(* CODESYS project maincontrol.library
   DefaultNamespace: KOSTAL.AF2024.Core.MainControl
   DocFormat: reStructuredText
   Description: Base Class of Machnie Main Control with 
      Cell_EXT using the ListOfInterface library instead of the generic array.
      The handler for the subscribers/stations is provided as well.
   Author: Frank Dümpelmann
   Title: KOSTAL.AF2024.Core.MainControl
   Version: 1.0.0.0
   Company: KOSTAL GmbH & Co.KG
   Placeholder: KOSTAL.AF2024.Core.MainControl

Project tree, tasks and I/O mapping:
  libraries: KOSTAL.AF2024.Core.functionResponse, 1.0.0.0 (KOSTAL GmbH & Co.KG); KOSTAL.AF2024.Core.ID, 1.0.0.0 (KOSTAL GmbH & Co.KG); KOSTAL.AF2024.Core.ListOf, 1.0.0.0 (KOSTAL GmbH & Co.KG); KOSTAL.AF2024.Core.Process, 1.0.0.0 (KOSTAL GmbH & Co.KG); KOSTAL.AF2024.Core.Settings, 1.0.0.0 (KOSTAL GmbH & Co.KG); KOSTAL.AF2024.Core.StringTools, 1.0.0.0 (KOSTAL GmbH & Co.KG); KOSTAL.AF2024.Core.System, 1.0.0.0 (KOSTAL GmbH & Co.KG)
  MainControl/
    Participant/
      ListOf/
        function block FB_ListOfParticipant [ST]: _setResult, _verifyMember, AddMember, Clear, Get_Member, IsValidParticipant, NumberOfMember, RegKey, RemoveMember, RemoveMemberByNumber
        interface I_ListOfParticipant: NumberOfMember, RegKey
        interface I_ListOfParticipant_Owner: AddMember, Clear, Get_Member, IsValidParticipant, NumberOfMember, RegKey, RemoveMember, RemoveMemberByNumber
      function block FB_Participant [ST]: FB_init, _clearRegisterInformation, Register, ParticipantName, Condition, Demand, ID, Linked, Mode, State
      interface I_Participant: Demand, ID, Mode, Register, Condition, ParticipantName, State, Linked
    function block FB_MainControl [ST]: _all_ErrorFree, _all_Finish, _all_Home, _all_OnToHome, _all_PowerOff, _all_PowerOn, _all_Run, _getNameAndID, _setResult, FB_exit, FB_init, Register, Unregister, condition, Demand, Device_ID, enableStopMode, ID, ID_RO, Mode, Participants, RunEmpty, step
    interface I_MainControl: condition, Demand, Device_ID, enableStopMode, ID_RO, Mode, Participants, RunEmpty, step
  MainControlState/
    interface I_T_MainControlState: CopyTo, Home, OnToHome, PowerOff, PowerOn, Run, RunToHome
    interface I_T_MainControlState_CopyFrom: CopyFrom
    interface I_T_MainControlState_Owner: clear, CopyFrom, CopyTo, Home, OnToHome, PowerOff, PowerOn, Run, RunToHome, SetUnique_Home, SetUnique_OnToHome, SetUnique_PowerOff, SetUnique_PowerOn, SetUnique_Run, SetUnique_RunToHome
    function block T_MainControlState [ST]: _clear_state, clear, CopyFrom, CopyTo, Home, OnToHome, PowerOff, PowerOn, Run, RunToHome, SetUnique_Home, SetUnique_OnToHome, SetUnique_PowerOff, SetUnique_PowerOn, SetUnique_Run, SetUnique_RunToHome
  ParticipantState/
    interface I_T_ParticipantState: Busy, CopyTo, Finish, Home, OnToHome, PowerOff, PowerOn
    interface I_T_ParticipantState_CopyFrom: CopyFrom
    interface I_T_ParticipantState_Owner: Busy, clear, CopyFrom, CopyTo, Finish, Home, OnToHome, PowerOff, PowerOn, SetUnique_Busy, SetUnique_Finish, SetUnique_Home, SetUnique_OnToHome, SetUnique_PowerOff, SetUnique_PowerOn
    function block T_ParticipantState [ST]: _clear_state, Busy, clear, CopyFrom, CopyTo, Finish, Home, OnToHome, PowerOff, PowerOn, SetUnique_Busy, SetUnique_Finish, SetUnique_Home, SetUnique_OnToHome, SetUnique_PowerOff, SetUnique_PowerOn
  Project Information/
    function F_GetCompany [ST]
    function F_GetTitle [ST]
    function F_GetVersion [ST]
  Version/
    global variables Global_Version
*)

// Version/Global_Version
{attribute 'TcGenerated'}
{attribute 'no-analysis'}
{attribute 'linkalways'}
// This function has been automatically generated from the project information.
VAR_GLOBAL CONSTANT
	{attribute 'const_non_replaced'}
	stLibVersion_KOSTAL_AF2024_Core_MainControl : ST_LibVersion := (iMajor := 1, iMinor := 0, iBuild := 0, iRevision := 0, nFlags := 0, sVersion := '1.0.0.0');
END_VAR

// MainControl/Participant/ListOf/FB_ListOfParticipant
(*
Extends the generic class with typed content.
*)
FUNCTION_BLOCK FB_ListOfParticipant EXTENDS KOSTAL_AF2024_Core_ListOf._FB_Interface_Base IMPLEMENTS I_ListOfParticipant, I_ListOfParticipant_Owner

VAR
	_PH_ID				: KOSTAL_AF2024_Core_ID.T_ID;	//placeholder for interfaces
	_PH_Condition 		: KOSTAL_AF2024_Core_Process.FB_processCondition;	//placeholder for interfaces
	_PH_State		 	: T_ParticipantState;	//placeholder for interfaces
	_PH_MainControlDemand		: T_MainControlState;	//placeholder for interfaces
	_PH_MainControlMode 		: KOSTAL_AF2024_Core_Process.T_processMode;	//placeholder for interfaces

	_Dummy	:	FB_Participant(ID:= _PH_ID, Condition:= _PH_Condition, State:= _PH_State);
END_VAR

METHOD PROTECTED _setResult
VAR_INPUT
	Status	: KOSTAL_AF2024_Core_Settings.T_MaxString;
	Success	: BOOL;
	Result	: KOSTAL_AF2024_Core_functionResponse.I_T_functionResponse_Owner;
END_VAR

IF Result = 0 THEN RETURN;	END_IF

Result.status:= Status;
Result.success:= Success;
END_METHOD

(*
	integrate here the veryfing of your interface type 
	only if verifing is passed [_verifyMember:= TRUE] the called metode will proceeded 
*)
METHOD PROTECTED _verifyMember : BOOL

VAR_INPUT
	Member	: KOSTAL_AF2024_Core_System.I_Interface;
	Result	: KOSTAL_AF2024_Core_functionResponse.I_T_functionResponse_Owner;
END_VAR

VAR
	_obj	: I_Participant;
	_bResult: BOOL;
END_VAR

_verifyMember:= SUPER^._verifyMember(Member, Result);

IF NOT _verifyMember THEN RETURN;	END_IF

//if member is I_participant?
_bResult:= __QUERYINTERFACE(Member, _obj);

IF NOT _bResult OR (_obj = 0) THEN
	IF Result <> 0 THEN
		Result.success:= FALSE;
		Result.status:= "no valid interface found";	
	END_IF	
	RETURN;
END_IF

//if 
IF NOT IsValidParticipant(_obj, Result)	THEN RETURN;	END_IF

_verifyMember:= TRUE;
END_METHOD

(*
	add new {Member} to end of list
*)
METHOD PUBLIC AddMember : BOOL

VAR_INPUT
	Member	: KOSTAL_AF2024_Core_System.I_Interface;
	Result	: KOSTAL_AF2024_Core_functionResponse.I_T_functionResponse_Owner;
END_VAR

AddMember:= SUPER^._addMember(Member, Result);

IF AddMember THEN	AddMember:= SUPER^._checkConsistency(Result);	END_IF
END_METHOD

//Clear the whole content
METHOD PUBLIC Clear

SUPER^._clear();
END_METHOD

METHOD PUBLIC Get_Member : I_Participant
VAR_INPUT
	Number		: UDINT;	//Participant which shall return
	Response	: KOSTAL_AF2024_Core_functionResponse.I_T_functionResponse_Owner;
END_VAR

VAR
	_Response	: KOSTAL_AF2024_Core_functionResponse.T_functionResponse;
	_Member			:	KOSTAL_AF2024_Core_System.I_Interface; 
	_obj			: I_Participant;
	_bResult	: BOOL;
	_found		: BOOL;
END_VAR
Get_Member:= _Dummy;

IF Number = 0 THEN
	IF Response <> 0 THEN	
		Response.success:= FALSE;	Response.status:= "Number is out of range";	
	END_IF
	RETURN;
END_IF

_found := _findMemberByIndex(Number - 1, _Member, _Response);
 
IF NOT _found OR NOT _Response.success THEN
 IF Response <> 0 THEN 
	Response.CopyFrom(_Response);	
	END_IF
 RETURN;
END_IF

_bResult:= __QUERYINTERFACE(_Member, _obj);

IF NOT _bResult THEN
	_Response.success:= FALSE;	_Response.status:= "__QUERYINTERFACE (I_RO) failed";
	IF Response <> 0 THEN 
		Response.CopyFrom(_Response);		
		END_IF
	RETURN;
END_IF

_Response.success:= TRUE;	_Response.status:= "Successful";
IF Response <> 0 THEN 
	Response.CopyFrom(_Response);	
END_IF

Get_Member:= _obj;
END_METHOD

METHOD PUBLIC IsValidParticipant : BOOL
VAR_INPUT
	Participant	: I_Participant;
	Result			: KOSTAL_AF2024_Core_functionResponse.I_T_functionResponse_Owner;
END_VAR

VAR
	_oParticipant 				: I_Participant;
	_bResult			: BOOL;
END_VAR
IsValidParticipant:= FALSE;

IF	Participant = 0 THEN	_setResult("no valid I_Participant INTERFACE", FALSE, Result);	RETURN; END_IF	

_bResult:= __QUERYINTERFACE( Participant, _oParticipant);

IF NOT _bResult 									THEN	_setResult("no valid I_Participant INTERFACE", FALSE, Result);	
ELSIF	_oParticipant = 0 									THEN	_setResult("no valid I_Participant INTERFACE", FALSE, Result);	
ELSIF	Participant = 0 						THEN	_setResult("no valid I_Participant INTERFACE", FALSE, Result);	
ELSIF Participant.Demand = 0	THEN	_setResult("no valid MainControlDemand INTERFACE", FALSE, Result);	
ELSIF Participant.Mode = 0		THEN	_setResult("no valid Mode INTERFACE", FALSE, Result);	
ELSIF Participant.Condition = 0		THEN	_setResult("no valid Condition INTERFACE", FALSE, Result);	
ELSIF Participant.ID = 0					THEN	_setResult("no valid ID INTERFACE", FALSE, Result);	
ELSIF Participant.State = 0				THEN	_setResult("no valid State INTERFACE", FALSE, Result);	
ELSE	IsValidParticipant:= TRUE;
END_IF
END_METHOD

//return the nnumber of items in List
PROPERTY PUBLIC NumberOfMember : UDINT
GET

NumberOfMember:= _NumberOfMember;
END_GET
END_PROPERTY

PROPERTY PUBLIC RegKey : UDINT
GET

RegKey:= _RegKey;
END_GET
END_PROPERTY

(*
	remove given {Member} from List
*)
METHOD PUBLIC RemoveMember : BOOL
VAR_INPUT
	Member	: KOSTAL_AF2024_Core_System.I_Interface;
	Result	: KOSTAL_AF2024_Core_functionResponse.I_T_functionResponse_Owner;
END_VAR

IF NOT _verifyMember(Member, Result) THEN	RETURN;	END_IF

RemoveMember:= _removeMember(Member, Result);

IF RemoveMember THEN	RemoveMember:= SUPER^._checkConsistency(Result);	END_IF
END_METHOD

(*
	remove given {Number} from List
*)
METHOD PUBLIC RemoveMemberByNumber : BOOL
VAR_INPUT
	Number	: UDINT;	//Position which shall deleted
	Result	: KOSTAL_AF2024_Core_functionResponse.I_T_functionResponse_Owner;
END_VAR
IF Number = 0 THEN
	IF Result <> 0  THEN
		Result.success:= FALSE;	
		Result.status:= "Number is out of range";	
	END_IF
	RETURN;
END_IF

RemoveMemberByNumber:= _removeMemberByIndex(Number - 1, Result);

IF RemoveMemberByNumber THEN	RemoveMemberByNumber:= SUPER^._checkConsistency(Result);	END_IF
END_METHOD

END_FUNCTION_BLOCK

// MainControl/Participant/ListOf/I_ListOfParticipant
(*
	Read-Only access to List
*)
INTERFACE I_ListOfParticipant EXTENDS KOSTAL_AF2024_Core_ListOf._I_Interface_Base

PROPERTY PUBLIC NumberOfMember : UDINT
GET
END_GET
END_PROPERTY

PROPERTY PUBLIC RegKey : UDINT
GET
END_GET
END_PROPERTY

END_INTERFACE

// MainControl/Participant/ListOf/I_ListOfParticipant_Owner
(*
	full access to List
*)
INTERFACE I_ListOfParticipant_Owner EXTENDS KOSTAL_AF2024_Core_ListOf._I_Interface_Base_Owner

(*
	add new {Member} to end of list
*)
METHOD PUBLIC AddMember : BOOL

VAR_INPUT
	Member	: KOSTAL_AF2024_Core_System.I_Interface;
	Result	: KOSTAL_AF2024_Core_functionResponse.I_T_functionResponse_Owner;
END_VAR
END_METHOD

//Clear the whole content
METHOD PUBLIC Clear
END_METHOD

METHOD PUBLIC Get_Member : I_Participant
VAR_INPUT
	Number		: UDINT;	//Participant which shall return
	Response	: KOSTAL_AF2024_Core_functionResponse.I_T_functionResponse_Owner;
END_VAR
END_METHOD

METHOD PUBLIC IsValidParticipant : BOOL
VAR_INPUT
	Participant	: I_Participant;
	Result			: KOSTAL_AF2024_Core_functionResponse.I_T_functionResponse_Owner;
END_VAR
END_METHOD

//return the nnumber of items in List
PROPERTY PUBLIC NumberOfMember : UDINT
GET
END_GET
END_PROPERTY

PROPERTY PUBLIC RegKey : UDINT
GET
END_GET
END_PROPERTY

(*
	remove given {Member} from List
*)
METHOD PUBLIC RemoveMember : BOOL
VAR_INPUT
	Member	: KOSTAL_AF2024_Core_System.I_Interface;
	Result	: KOSTAL_AF2024_Core_functionResponse.I_T_functionResponse_Owner;
END_VAR
END_METHOD

(*
	remove given {Number} from List
*)
METHOD PUBLIC RemoveMemberByNumber : BOOL
VAR_INPUT
	Number	: UDINT;	//Position which shall deleted
	Result	: KOSTAL_AF2024_Core_functionResponse.I_T_functionResponse_Owner;
END_VAR
END_METHOD

END_INTERFACE

// MainControl/Participant/I_Participant
(*

:Author: Frank Dümpelmann <f.duempelmann@kostal.com>, Martin Hundt <m.hundt@kostal.com>
:Date: 2018-10-29

Function
========
Interface for communication between stations and MainControl

Usage notes
===============
| All stations must be implemented with this interface



*)

INTERFACE I_Participant EXTENDS KOSTAL_AF2024_Core_System.I_Interface

(*State requirement for the participant*)
PROPERTY Demand : I_T_MainControlState
GET
END_GET
END_PROPERTY

(*
	ID of the participant
	{name} will handeld by participant
	{key} will handled by MainControl. 
*)
PROPERTY ID : KOSTAL_AF2024_Core_ID.I_T_ID
GET
END_GET
END_PROPERTY

(*Mode information for the participant*)
PROPERTY Mode : KOSTAL_AF2024_Core_process.I_T_processMode
GET
END_GET
END_PROPERTY

(*
	Called by MainControl
*)
METHOD PUBLIC Register
VAR_INPUT
	MainControlDemand	: I_T_MainControlState;
	MainControlMode		: KOSTAL_AF2024_Core_process.I_T_processMode;
	RegKey			: UDINT;
	Linked			: BOOL;
END_VAR
END_METHOD

(*Condition of the participant*)
PROPERTY Condition : KOSTAL_AF2024_Core_process.I_processCondition
GET
END_GET
END_PROPERTY

PROPERTY PUBLIC ParticipantName : KOSTAL_AF2024_Core_Settings.T_MaxString
GET
END_GET
END_PROPERTY

(*State of the participant*)
PROPERTY State : I_T_ParticipantState
GET
END_GET
END_PROPERTY

PROPERTY PUBLIC Linked : BOOL
GET
END_GET
END_PROPERTY

END_INTERFACE

// MainControlState/I_T_MainControlState
INTERFACE I_T_MainControlState EXTENDS KOSTAL_AF2024_Core_System.I_Interface

METHOD PUBLIC CopyTo
VAR_INPUT
	IN	:	I_T_MainControlState_CopyFrom;
END_VAR
END_METHOD

PROPERTY PUBLIC Home : BOOL
GET
END_GET
END_PROPERTY

PROPERTY PUBLIC OnToHome : BOOL
GET
END_GET
END_PROPERTY

PROPERTY PUBLIC PowerOff : BOOL
GET
END_GET
END_PROPERTY

PROPERTY PUBLIC PowerOn : BOOL
GET
END_GET
END_PROPERTY

PROPERTY PUBLIC Run : BOOL
GET
END_GET
END_PROPERTY

PROPERTY PUBLIC RunToHome : BOOL
GET
END_GET
END_PROPERTY

END_INTERFACE

// MainControlState/I_T_MainControlState_CopyFrom
INTERFACE I_T_MainControlState_CopyFrom EXTENDS KOSTAL_AF2024_Core_System.I_Interface

METHOD PUBLIC CopyFrom
VAR_INPUT
	IN	: I_T_MainControlState;
END_VAR
END_METHOD

END_INTERFACE

// ParticipantState/I_T_ParticipantState
INTERFACE I_T_ParticipantState EXTENDS KOSTAL_AF2024_Core_System.I_Interface

PROPERTY PUBLIC Busy : BOOL
GET
END_GET
END_PROPERTY

METHOD PUBLIC CopyTo
VAR_INPUT
	IN	:	I_T_ParticipantState_CopyFrom;
END_VAR
END_METHOD

PROPERTY PUBLIC Finish : BOOL
GET
END_GET
END_PROPERTY

PROPERTY PUBLIC Home : BOOL
GET
END_GET
END_PROPERTY

PROPERTY PUBLIC OnToHome : BOOL
GET
END_GET
END_PROPERTY

PROPERTY PUBLIC PowerOff : BOOL
GET
END_GET
END_PROPERTY

PROPERTY PUBLIC PowerOn : BOOL
GET
END_GET
END_PROPERTY

END_INTERFACE

// ParticipantState/I_T_ParticipantState_CopyFrom
INTERFACE I_T_ParticipantState_CopyFrom EXTENDS KOSTAL_AF2024_Core_System.I_Interface

METHOD PUBLIC CopyFrom
VAR_INPUT
	IN	: I_T_ParticipantState;
END_VAR
END_METHOD

END_INTERFACE

// ParticipantState/T_ParticipantState
(*

:Author: Martin Hundt <m.hundt@kostal.com>
:Date: 2024-01-31

Function
========
Data type representing the process state of a Main Control's participant

Methods and Properties
======================
| Properties represent the possible process states 
| Methods setUnique_... set the corresponding state and clear the others
| Alternatively, states can be set independent of the others using the properties 
| Methods starting with an underline(_) are internally used and can be ignored by the user
*)
{attribute 'enable_dynamic_creation'}
FUNCTION_BLOCK PUBLIC T_ParticipantState IMPLEMENTS I_T_ParticipantState, I_T_ParticipantState_CopyFrom, I_T_ParticipantState_Owner

VAR
	_powerOff 		: BOOL;	//BOOL
	_powerOn 		: BOOL;	//BOOL
	_onToHome 		: BOOL;	//BOOL
	_home 			: BOOL;	//BOOL
	_busy 			: BOOL;	//BOOL
	_finish 		: BOOL;	//BOOL
END_VAR

METHOD PROTECTED _clear_state

_busy		:= FALSE;
_onToHome	:= FALSE;
_finish		:= FALSE;
_powerOff		:= FALSE;
_powerOn			:= FALSE;
_home		:= FALSE;
END_METHOD

PROPERTY PUBLIC Busy : BOOL
GET

Busy:= _busy;
END_GET
SET

_busy:= Busy;
END_SET
END_PROPERTY

METHOD PUBLIC clear

_clear_state();
END_METHOD

METHOD PUBLIC CopyFrom
VAR_INPUT
	IN	: I_T_ParticipantState;
END_VAR

IF IN = 0 THEN	RETURN;	END_IF

_powerOff				:= IN.PowerOff;
_powerOn					:= IN.PowerOn;
_onToHome	:= IN.OnToHome;
_busy				:= IN.Busy;
_home			:= IN.Home;
_finish			:= IN.Finish;
END_METHOD

METHOD PUBLIC CopyTo
VAR_INPUT
	IN	:	I_T_ParticipantState_CopyFrom;
END_VAR

IF IN = 0 THEN	RETURN;	END_IF

IN.CopyFrom(THIS^);
END_METHOD

PROPERTY PUBLIC Finish : BOOL
GET

Finish:= _finish;
END_GET
SET

_finish:= Finish;
END_SET
END_PROPERTY

PROPERTY PUBLIC Home : BOOL
GET

Home:= _home;
END_GET
SET

_home:= Home;
END_SET
END_PROPERTY

PROPERTY PUBLIC OnToHome : BOOL
GET

OnToHome:= _onToHome;
END_GET
SET

_onToHome:= OnToHome;
END_SET
END_PROPERTY

PROPERTY PUBLIC PowerOff : BOOL
GET

PowerOff:= _powerOff;
END_GET
SET

_powerOff:= PowerOff;
END_SET
END_PROPERTY

PROPERTY PUBLIC PowerOn : BOOL
GET

PowerOn:= _powerOn;
END_GET
SET

_powerOn:= PowerOn;
END_SET
END_PROPERTY

METHOD PUBLIC SetUnique_Busy

_clear_state();

_busy:= TRUE;
END_METHOD

METHOD PUBLIC SetUnique_Finish

_clear_state();

_finish:= TRUE;
END_METHOD

METHOD PUBLIC SetUnique_Home

_clear_state();

_home:= TRUE;
END_METHOD

METHOD PUBLIC SetUnique_OnToHome

_clear_state();

_onToHome:= TRUE;
END_METHOD

METHOD PUBLIC SetUnique_PowerOff

_clear_state();

_powerOff:= TRUE;
END_METHOD

METHOD PUBLIC SetUnique_PowerOn

_clear_state();

_powerOn:= TRUE;
END_METHOD

END_FUNCTION_BLOCK

// ParticipantState/I_T_ParticipantState_Owner
INTERFACE I_T_ParticipantState_Owner EXTENDS KOSTAL_AF2024_Core_System.I_Interface

PROPERTY PUBLIC Busy : BOOL
GET
END_GET
SET
END_SET
END_PROPERTY

METHOD PUBLIC clear
END_METHOD

METHOD PUBLIC CopyFrom
VAR_INPUT
	IN	: I_T_ParticipantState;
END_VAR
END_METHOD

METHOD PUBLIC CopyTo
VAR_INPUT
	IN	:	I_T_ParticipantState_CopyFrom;
END_VAR
END_METHOD

PROPERTY PUBLIC Finish : BOOL
GET
END_GET
SET
END_SET
END_PROPERTY

PROPERTY PUBLIC Home : BOOL
GET
END_GET
SET
END_SET
END_PROPERTY

PROPERTY PUBLIC OnToHome : BOOL
GET
END_GET
SET
END_SET
END_PROPERTY

PROPERTY PUBLIC PowerOff : BOOL
GET
END_GET
SET
END_SET
END_PROPERTY

PROPERTY PUBLIC PowerOn : BOOL
GET
END_GET
SET
END_SET
END_PROPERTY

METHOD PUBLIC SetUnique_Busy
END_METHOD

METHOD PUBLIC SetUnique_Finish
END_METHOD

METHOD PUBLIC SetUnique_Home
END_METHOD

METHOD PUBLIC SetUnique_OnToHome
END_METHOD

METHOD PUBLIC SetUnique_PowerOff
END_METHOD

METHOD PUBLIC SetUnique_PowerOn
END_METHOD

END_INTERFACE

// MainControlState/T_MainControlState
(*

:Author: Martin Hundt <m.hundt@kostal.com>
:Date: 2024-01-31

Function
========
Data type representing the process state of the Main Control

Methods and Properties
======================
| Properties represent the possible process states 
| Methods setUnique_... set the corresponding state and clear the others
| Alternatively, states can be set independent of the others using the properties 
| Methods starting with an underline(_) are internally used and can be ignored by the user
*)
{attribute 'enable_dynamic_creation'}
FUNCTION_BLOCK PUBLIC T_MainControlState IMPLEMENTS I_T_MainControlState, I_T_MainControlState_CopyFrom, I_T_MainControlState_Owner

VAR
	_powerOff 			: BOOL;	//BOOL
	_powerOn 			: BOOL;	//BOOL
	_onToHome 		: BOOL;	//BOOL
	_home 			: BOOL;	//BOOL
	_run 			: BOOL;	//BOOL
	_runToHome 		: BOOL;	//BOOL
END_VAR

METHOD PROTECTED _clear_state

_run		:= FALSE;
_onToHome	:= FALSE;
_runToHome		:= FALSE;
_powerOff		:= FALSE;
_powerOn			:= FALSE;
_home		:= FALSE;
END_METHOD

METHOD PUBLIC clear

_clear_state();
END_METHOD

METHOD PUBLIC CopyFrom
VAR_INPUT
	IN	: I_T_MainControlState;
END_VAR

IF IN = 0 THEN	RETURN;	END_IF

_powerOff				:= IN.PowerOff;
_powerOn					:= IN.PowerOn;
_onToHome	:= IN.OnToHome;
_run				:= IN.Run;
_home			:= IN.Home;
_runToHome			:= IN.RunToHome;
END_METHOD

METHOD PUBLIC CopyTo
VAR_INPUT
	IN	:	I_T_MainControlState_CopyFrom;
END_VAR

IF IN = 0 THEN	RETURN;	END_IF

IN.CopyFrom(THIS^);
END_METHOD

PROPERTY PUBLIC Home : BOOL
GET

Home:= _home;
END_GET
SET

_home:= Home;
END_SET
END_PROPERTY

PROPERTY PUBLIC OnToHome : BOOL
GET

OnToHome:= _onToHome;
END_GET
SET

_onToHome:= OnToHome;
END_SET
END_PROPERTY

PROPERTY PUBLIC PowerOff : BOOL
GET

PowerOff:= _powerOff;
END_GET
SET

_powerOff:= PowerOff;
END_SET
END_PROPERTY

PROPERTY PUBLIC PowerOn : BOOL
GET

PowerOn:= _powerOn;
END_GET
SET

_powerOn:= PowerOn;
END_SET
END_PROPERTY

PROPERTY PUBLIC Run : BOOL
GET

Run:= _run;
END_GET
SET

_run:= Run;
END_SET
END_PROPERTY

PROPERTY PUBLIC RunToHome : BOOL
GET

RunToHome:= _runToHome;
END_GET
SET

_runToHome:= RunToHome;
END_SET
END_PROPERTY

METHOD PUBLIC SetUnique_Home

_clear_state();

_home:= TRUE;
END_METHOD

METHOD PUBLIC SetUnique_OnToHome

_clear_state();

_onToHome:= TRUE;
END_METHOD

METHOD PUBLIC SetUnique_PowerOff

_clear_state();

_powerOff:= TRUE;
END_METHOD

METHOD PUBLIC SetUnique_PowerOn

_clear_state();

_powerOn:= TRUE;
END_METHOD

METHOD PUBLIC SetUnique_Run

_clear_state();

_run:= TRUE;
END_METHOD

METHOD PUBLIC SetUnique_RunToHome

_clear_state();

_runToHome:= TRUE;
END_METHOD

END_FUNCTION_BLOCK

// MainControlState/I_T_MainControlState_Owner
INTERFACE I_T_MainControlState_Owner EXTENDS KOSTAL_AF2024_Core_System.I_Interface

METHOD PUBLIC clear
END_METHOD

METHOD PUBLIC CopyFrom
VAR_INPUT
	IN	: I_T_MainControlState;
END_VAR
END_METHOD

METHOD PUBLIC CopyTo
VAR_INPUT
	IN	:	I_T_MainControlState_CopyFrom;
END_VAR
END_METHOD

PROPERTY PUBLIC Home : BOOL
GET
END_GET
SET
END_SET
END_PROPERTY

PROPERTY PUBLIC OnToHome : BOOL
GET
END_GET
SET
END_SET
END_PROPERTY

PROPERTY PUBLIC PowerOff : BOOL
GET
END_GET
SET
END_SET
END_PROPERTY

PROPERTY PUBLIC PowerOn : BOOL
GET
END_GET
SET
END_SET
END_PROPERTY

PROPERTY PUBLIC Run : BOOL
GET
END_GET
SET
END_SET
END_PROPERTY

PROPERTY PUBLIC RunToHome : BOOL
GET
END_GET
SET
END_SET
END_PROPERTY

METHOD PUBLIC SetUnique_Home
END_METHOD

METHOD PUBLIC SetUnique_OnToHome
END_METHOD

METHOD PUBLIC SetUnique_PowerOff
END_METHOD

METHOD PUBLIC SetUnique_PowerOn
END_METHOD

METHOD PUBLIC SetUnique_Run
END_METHOD

METHOD PUBLIC SetUnique_RunToHome
END_METHOD

END_INTERFACE

// MainControl/Participant/FB_Participant
(*
	Use in Participants to handle the I_MainControl interface
*)
FUNCTION_BLOCK PUBLIC FB_Participant IMPLEMENTS I_Participant

VAR
	{region 'placeholder for interfaces'}
		_PH_ID				: KOSTAL_AF2024_Core_ID.T_ID;	//placeholder for interfaces
		_PH_Condition 	: KOSTAL_AF2024_Core_process.FB_processCondition;	//placeholder for interfaces
		_PH_State		: T_ParticipantState;	//placeholder for interfaces
		_PH_MainControlDemand 	: T_MainControlState;	//placeholder for interfaces
		_PH_Mode 	: KOSTAL_AF2024_Core_process.T_processMode;	//placeholder for interfaces
	{endregion}

	_IID						: KOSTAL_AF2024_Core_ID.I_T_ID;
	_ICondition 	: KOSTAL_AF2024_Core_process.I_processCondition;
	_IState		 	: I_T_ParticipantState;
	_IMainControlDemand	: I_T_MainControlState;
	_IMainControlMode 		: KOSTAL_AF2024_Core_process.I_T_processMode;
	
	//{Name} FROM participant
	_ParticipantName	: KOSTAL_AF2024_Core_Settings.T_MaxString;
	_RegKey	: UDINT;
	_Linked	: BOOL;
	
END_VAR

METHOD FB_init : BOOL
VAR_INPUT
	bInitRetains : BOOL; // if TRUE, the retain variables are initialized (warm start / cold start)
	bInCopyCode : BOOL;  // if TRUE, the instance afterwards gets moved into the copy code (online change)

	ID					:	KOSTAL_AF2024_Core_ID.I_T_ID;
	Condition		: KOSTAL_AF2024_Core_Process.I_processCondition;
	State				: I_T_ParticipantState;
END_VAR

VAR
	_bResult			: BOOL;
	_oID					:	KOSTAL_AF2024_Core_ID.I_T_ID;
	_oCondition		: KOSTAL_AF2024_Core_Process.I_processCondition;
	_oState				: I_T_ParticipantState;
END_VAR

_PH_ID.clear();
_PH_Condition.clear();
_PH_State.clear();

_PH_MainControlDemand.clear();	
_IMainControlDemand:= _PH_MainControlDemand;

_PH_Mode.clear();		
_IMainControlMode	:= _PH_Mode;		

_bResult:= __QUERYINTERFACE(ID, _oID);
IF _bResult AND (_oID <> 0) THEN	
	_IID	:= ID;
ELSE															
	_IID	:= _PH_ID;
END_IF

_bResult:= __QUERYINTERFACE(Condition, _oCondition);
IF _bResult AND (_oCondition <> 0) THEN	
	_ICondition	:= Condition;
ELSE																		
	_ICondition	:= _PH_Condition;
END_IF

_bResult:= __QUERYINTERFACE(State, _oState);
IF _bResult AND (_oState <> 0) THEN	
	_IState	:= State;
ELSE																
	_IState	:= _PH_State;
END_IF

_RegKey:= 0;
_Linked:= FALSE;
END_METHOD

METHOD PROTECTED _clearRegisterInformation

_IMainControlDemand	:= _PH_MainControlDemand;
_IMainControlMode 		:= _PH_Mode;
END_METHOD

(*
	Called by MainControl
*)
METHOD PUBLIC Register
VAR_INPUT
	MainControlDemand	: I_T_MainControlState;
	MainControlMode		: KOSTAL_AF2024_Core_process.I_T_processMode;

	RegKey			: UDINT;
	Linked			: BOOL;
END_VAR

VAR
	_oMainControlMode 		: KOSTAL_AF2024_Core_process.I_T_processMode;
	_oMainControlDemand	: I_T_MainControlState;
	_oID					: KOSTAL_AF2024_Core_ID.I_T_ID;
	_bResult: BOOL;
END_VAR
_Linked:= Linked;
_RegKey:= RegKey;


IF NOT _Linked THEN	_clearRegisterInformation();	

ELSE

	_bResult:= __QUERYINTERFACE(MainControlDemand, _oMainControlDemand);
	IF _bResult AND (_oMainControlDemand <> 0) THEN	_IMainControlDemand:= MainControlDemand;	
	ELSE																			_IMainControlDemand:= _PH_MainControlDemand;	
	END_IF
	
	_bResult:= __QUERYINTERFACE(MainControlMode, _oMainControlMode);
	IF _bResult AND (_oMainControlMode <> 0) THEN	_IMainControlMode:= MainControlMode;	
	ELSE																		_IMainControlMode:= _PH_Mode;	
	END_IF
	


END_IF
END_METHOD

PROPERTY PUBLIC ParticipantName : KOSTAL_AF2024_Core_Settings.T_MaxString
GET

ParticipantName:= _ParticipantName;
END_GET
SET

_ParticipantName:= ParticipantName;
END_SET
END_PROPERTY

(*Condition of the participant*)
PROPERTY Condition : KOSTAL_AF2024_Core_process.I_processCondition
GET

Condition:= _ICondition;
END_GET
END_PROPERTY

(*State requirement for the participant*)
PROPERTY Demand : I_T_MainControlState
GET

Demand:= _IMainControlDemand;
END_GET
END_PROPERTY

(*ID of the participant*)
PROPERTY ID : KOSTAL_AF2024_Core_ID.I_T_ID
GET

ID:= _IID;
END_GET
END_PROPERTY

PROPERTY PUBLIC Linked : BOOL
GET

Linked:= _Linked;
END_GET
END_PROPERTY

(*Mode information for the participant*)
PROPERTY Mode : KOSTAL_AF2024_Core_process.I_T_processMode
GET

Mode:= _IMainControlMode;
END_GET
END_PROPERTY

(*State of the participant*)
PROPERTY State : I_T_ParticipantState
GET

State:= _IState;
END_GET
END_PROPERTY

END_FUNCTION_BLOCK

// MainControl/I_MainControl
INTERFACE I_MainControl EXTENDS KOSTAL_AF2024_Core_System.I_Interface

PROPERTY PUBLIC condition : KOSTAL_AF2024_Core_process.I_processCondition
GET
END_GET
END_PROPERTY

PROPERTY PUBLIC Demand : I_T_MainControlState
GET
END_GET
END_PROPERTY

PROPERTY PUBLIC Device_ID : KOSTAL_AF2024_Core_Settings.T_MaxString
GET
END_GET
END_PROPERTY

PROPERTY PUBLIC enableStopMode : BOOL
GET
END_GET
END_PROPERTY

PROPERTY PUBLIC ID_RO : KOSTAL_AF2024_Core_ID.I_T_ID
GET
END_GET
END_PROPERTY

PROPERTY PUBLIC Mode : KOSTAL_AF2024_Core_process.I_T_processMode
GET
END_GET
END_PROPERTY

PROPERTY PUBLIC Participants : I_ListOfParticipant
GET
END_GET
END_PROPERTY

PROPERTY PUBLIC RunEmpty : BOOL
GET
END_GET
END_PROPERTY

PROPERTY PUBLIC step : KOSTAL_AF2024_Core_process.I_processStep
GET
END_GET
END_PROPERTY

END_INTERFACE

// MainControl/FB_MainControl
(*

:Author: Frank Dümpelmann <f.duempelmann@kostal.com>, Martin Hundt <m.hundt@kostal.com>
:Date: 2018-10-29

Function
========
Base class representing a machine's main control

Usage notes
===============
| Extend the base class to implement a main control

Methods and Properties
======================
| See best practice and project tempates

*)

FUNCTION_BLOCK PUBLIC FB_MainControl IMPLEMENTS I_MainControl
VAR
	

	_Participants	: FB_ListOfParticipant;
	
	_demand		: T_MainControlState;

	//my own
	_ID					: KOSTAL_AF2024_Core_ID.T_ID;
	//_state				: T_MainControlState;
	_condition	: KOSTAL_AF2024_Core_process.FB_ProcessCondition;
	_mode		: KOSTAL_AF2024_Core_process.T_processMode;


	_Device_ID	: KOSTAL_AF2024_Core_Settings.T_MaxString;		//PC name / name Function unit / controller name
	_runEmpty	: BOOL;
	_enableStopMode	: BOOL:= TRUE;

	_step					: KOSTAL_AF2024_Core_process.FB_processStep;	//Step Chain

END_VAR

(*
Description
===========
| Returns true when no stations in the MainControl has an error
*)
METHOD PROTECTED _all_ErrorFree : BOOL

VAR_INPUT
	Participant	: REFERENCE TO KOSTAL_AF2024_Core_Settings.T_MaxString;
END_VAR

VAR
	_udi				: UDINT;
	_Result			: KOSTAL_AF2024_Core_functionResponse.T_functionResponse;
	_Participant: I_Participant;
END_VAR
_all_ErrorFree:= FALSE;

IF __ISVALIDREF(Participant) THEN Participant:= "";	END_IF

FOR _udi:= 1 TO _Participants.NumberOfMember DO

	_Participant:= _Participants.Get_Member(_udi, _Result);

	IF _Participants.IsValidParticipant(_Participant, 0) AND _Result.success THEN
		IF NOT _Participant.Linked THEN	;	
		ELSIF _Participant.Condition.isError() THEN	
			IF __ISVALIDREF(Participant) THEN Participant:= _getNameAndID(_Participant);	END_IF
			RETURN;	
		END_IF
	END_IF

END_FOR

_all_ErrorFree:= TRUE;
END_METHOD

(*
Description
===========
| Returns true when all stations in the MainControl are finished
*)
METHOD PROTECTED _all_Finish : BOOL

VAR_INPUT
	Participant	: REFERENCE TO KOSTAL_AF2024_Core_Settings.T_MaxString;
END_VAR

VAR
	_udi				: UDINT;
	_Result			: KOSTAL_AF2024_Core_functionResponse.T_functionResponse;
	_Participant: I_Participant;
END_VAR
_all_FINISH:= FALSE;

IF __ISVALIDREF(Participant) THEN Participant:= "";	END_IF

FOR _udi:= 1 TO _Participants.NumberOfMember DO

	_Participant:= _Participants.Get_Member(_udi, _Result);

	IF _Participants.IsValidParticipant(_Participant, 0) AND _Result.success THEN
		IF NOT _Participant.Linked THEN	;	
		ELSIF NOT _Participant.State.Finish THEN	
			IF __ISVALIDREF(Participant) THEN Participant:= _getNameAndID(_Participant);	END_IF
			RETURN;	
		END_IF
	END_IF

END_FOR

_all_FINISH:= TRUE;
END_METHOD

(*
Description
===========
| Returns true when all stations in the MainControl are home
*)
METHOD PROTECTED _all_Home : BOOL

VAR_INPUT
	Participant	: REFERENCE TO KOSTAL_AF2024_Core_Settings.T_MaxString;
END_VAR

VAR
	_udi				: UDINT;
	_Result			: KOSTAL_AF2024_Core_functionResponse.T_functionResponse;
	_Participant: I_Participant;
END_VAR
_all_Home:= FALSE;

IF __ISVALIDREF(Participant) THEN Participant:= "";	END_IF

FOR _udi:= 1 TO _Participants.NumberOfMember DO

	_Participant:= _Participants.Get_Member(_udi, _Result);

	IF _Participants.IsValidParticipant(_Participant, 0) AND _Result.success THEN
		IF NOT _Participant.Linked THEN	;	
		ELSIF NOT _Participant.State.Home THEN
			IF __ISVALIDREF(Participant) THEN Participant:= _getNameAndID(_Participant);	END_IF
			RETURN;	
		END_IF
	END_IF

END_FOR


_all_Home:= TRUE;
END_METHOD

(*
Description
===========
| Returns true when all stations in the MainControl are in OnToHome state
*)
METHOD PROTECTED _all_OnToHome : BOOL

VAR_INPUT
	Participant	: REFERENCE TO KOSTAL_AF2024_Core_Settings.T_MaxString;
END_VAR

VAR
	_udi				: UDINT;
	_Result			: KOSTAL_AF2024_Core_functionResponse.T_functionResponse;
	_Participant: I_Participant;
END_VAR
_all_OnToHome:= FALSE;

IF __ISVALIDREF(Participant) THEN Participant:= "";	END_IF

FOR _udi:= 1 TO _Participants.NumberOfMember DO

	_Participant:= _Participants.Get_Member(_udi, _Result);

	IF _Participants.IsValidParticipant(_Participant, 0) AND _Result.success THEN
		IF NOT _Participant.Linked THEN	;	
		ELSIF NOT _Participant.State.OnToHome THEN	
			IF __ISVALIDREF(Participant) THEN Participant:= _getNameAndID(_Participant);	END_IF
			RETURN;	
		END_IF
	END_IF

END_FOR

_all_OnToHome:= TRUE;
END_METHOD

(*
Description
===========
| Returns true when all stations in the MainControl are off
*)
METHOD PROTECTED _all_PowerOff : BOOL

VAR_INPUT
	Participant	: REFERENCE TO KOSTAL_AF2024_Core_Settings.T_MaxString;
END_VAR

VAR
	_udi				: UDINT;
	_Result			: KOSTAL_AF2024_Core_functionResponse.T_functionResponse;
	_Participant: I_Participant;
END_VAR
_all_PowerOff:= FALSE;

IF __ISVALIDREF(Participant) THEN Participant:= "";	END_IF

FOR _udi:= 1 TO _Participants.NumberOfMember DO

	_Participant:= _Participants.Get_Member(_udi, _Result);

	IF _Participants.IsValidParticipant(_Participant, 0) AND _Result.success THEN
		IF NOT _Participant.Linked THEN	;	
		ELSIF NOT _Participant.State.PowerOff THEN	
			IF __ISVALIDREF(Participant) THEN Participant:= _getNameAndID(_Participant);	END_IF
			RETURN;	
		END_IF
	END_IF

END_FOR

_all_PowerOff:= TRUE;
END_METHOD

(*
Description
===========
| Returns true when all stations in the MainControl are on
*)
METHOD PROTECTED _all_PowerOn : BOOL


VAR_INPUT
	Participant	: REFERENCE TO KOSTAL_AF2024_Core_Settings.T_MaxString;
END_VAR

VAR
	_udi				: UDINT;
	_Result			: KOSTAL_AF2024_Core_functionResponse.T_functionResponse;
	_Participant: I_Participant;
END_VAR
_all_PowerOn:= FALSE;

IF __ISVALIDREF(Participant) THEN Participant:= "";	END_IF

FOR _udi:= 1 TO _Participants.NumberOfMember DO

	_Participant:= _Participants.Get_Member(_udi, _Result);

	IF _Participants.IsValidParticipant(_Participant, 0) AND _Result.success THEN
		IF NOT _Participant.Linked THEN	;	
		ELSIF NOT _Participant.State.PowerOn THEN	
			IF __ISVALIDREF(Participant) THEN Participant:= _getNameAndID(_Participant);	END_IF
			RETURN;	
		END_IF
	END_IF
		
END_FOR

_all_PowerOn:= TRUE;
END_METHOD

(*
Description
===========
| Returns true when all stations in the MainControl are in run state
*)
METHOD PROTECTED _all_Run : BOOL

VAR_INPUT
	Participant	: REFERENCE TO KOSTAL_AF2024_Core_Settings.T_MaxString;
END_VAR

VAR
	_udi				: UDINT;
	_Result			: KOSTAL_AF2024_Core_functionResponse.T_functionResponse;
	_Participant: I_Participant;
END_VAR
_all_RUN:= FALSE;

IF __ISVALIDREF(Participant) THEN Participant:= "";	END_IF

FOR _udi:= 1 TO _Participants.NumberOfMember DO

	_Participant:= _Participants.Get_Member(_udi, _Result);

	IF _Participants.IsValidParticipant(_Participant, 0) AND _Result.success THEN
		IF NOT _Participant.Linked THEN	;	
		ELSIF NOT _Participant.State.Busy THEN	
			IF __ISVALIDREF(Participant) THEN Participant:= _getNameAndID(_Participant);	END_IF
			RETURN;	
		END_IF
	END_IF
		
END_FOR

_all_RUN:= TRUE;
END_METHOD

METHOD PROTECTED _getNameAndID : KOSTAL_AF2024_Core_Settings.T_MaxString
VAR_INPUT
	_Participant	: I_Participant;
END_VAR

VAR
	_c	: Kostal_AF2024_Core_StringTools.FB_Concat;
END_VAR

IF _Participant = 0 THEN RETURN;	END_IF

_c.Clear();
_c.addContent(_Participant.ParticipantName);
_c.addContent("[");
_c.addContent(_Participant.ID.name);
_c.addContent("(");
_c.addContent(DINT_TO_WSTRING(_Participant.ID.key));
_c.addContent(")");
_c.addContent("]");
_getNameAndID:= _c.getResult();
_c.Clear();
END_METHOD

METHOD PROTECTED _setResult
VAR_INPUT
	Status	: KOSTAL_AF2024_Core_Settings.T_MaxString;
	Success	: BOOL;
	Result	: KOSTAL_AF2024_Core_functionResponse.I_T_functionResponse_Owner;
END_VAR

IF Result = 0 THEN RETURN;	END_IF

Result.status:= Status;
Result.success:= Success;
END_METHOD

METHOD FB_exit : BOOL
VAR_INPUT
	bInCopyCode : BOOL; // if TRUE, the exit method is called for exiting an instance that is copied afterwards (online change).
END_VAR

_Participants.Clear();
END_METHOD

METHOD FB_init : BOOL
VAR_INPUT
	bInitRetains 		: BOOL; // if TRUE, the retain variables are initialized (warm start / cold start)
	bInCopyCode 		: BOOL;  // if TRUE, the instance afterwards gets moved into the copy code (online change)
	EnableStopMode	: BOOL;
END_VAR

VAR
	_index: INT;	//INT
END_VAR

_Participants.Clear();

_enableStopMode				:= EnableStopMode;

_step.init();
END_METHOD

(*
Description
===========
| Adds a user to the link table at given position
| Parameters:
| 	component: user to be added
| 	index: position in link table

*)

METHOD PUBLIC Register : BOOL
VAR_INPUT
	Participant		: I_Participant;
	Result			: KOSTAL_AF2024_Core_functionResponse.I_T_functionResponse_Owner;
END_VAR

VAR
	_Result	: KOSTAL_AF2024_Core_functionResponse.T_functionResponse;
	//_ID	: KOSTAL_AF2024_Core_ID.FB_ID;
END_VAR

Register:= FALSE;

IF NOT _Participants.IsValidParticipant(Participant, Result) THEN	RETURN;	END_IF

  	
IF NOT _Participants.AddMember(Participant, _Result)	THEN
	_setResult(_Result.status, FALSE, Result);	RETURN;
END_IF


Participant.Register(MainControlDemand:= _demand, MainControlMode:= _mode, RegKey:= _Participants.RegKey, TRUE);

_setResult("Successful", TRUE, Result);	

Register:= TRUE;
END_METHOD

(*
Description
===========
| Adds a user to the link table at given position
| Parameters:
| 	component: user to be added
| 	index: position in link table

*)

METHOD PUBLIC Unregister : BOOL
VAR_INPUT
	Participant	: I_Participant;
	Result			: KOSTAL_AF2024_Core_functionResponse.I_T_functionResponse_Owner;
END_VAR

VAR
	_Result	: KOSTAL_AF2024_Core_functionResponse.T_functionResponse;
	_ID	: KOSTAL_AF2024_Core_ID.T_ID;
END_VAR
Unregister:= FALSE;

IF NOT _Participants.IsValidParticipant(Participant, Result) THEN	RETURN;	END_IF

  	
IF NOT _Participants.RemoveMember(Participant, _Result)	THEN
	_setResult(_Result.status, FALSE, Result);	RETURN;
END_IF

_ID.name:= "";
_ID.key:= 0;

Participant.Register(MainControlDemand:= 0, MainControlMode:= 0, RegKey:= UDINT#0, FALSE);

_setResult("Successful", TRUE, Result);	

Unregister:= TRUE;
END_METHOD

PROPERTY PUBLIC condition : KOSTAL_AF2024_Core_process.I_processCondition
GET

condition:= _condition;
END_GET
END_PROPERTY

PROPERTY PUBLIC Demand : I_T_MainControlState
GET

Demand:= _demand;
END_GET
END_PROPERTY

PROPERTY PUBLIC Device_ID : KOSTAL_AF2024_Core_Settings.T_MaxString
GET

Device_ID:= _Device_ID;
END_GET
SET

_Device_ID:= Device_ID;
END_SET
END_PROPERTY

PROPERTY PUBLIC enableStopMode : BOOL
GET

enableStopMode:= _enableStopMode;
END_GET
END_PROPERTY

PROPERTY PUBLIC ID : KOSTAL_AF2024_Core_ID.I_T_ID_Owner
GET

ID:= _ID;
END_GET
END_PROPERTY

PROPERTY PUBLIC ID_RO : KOSTAL_AF2024_Core_ID.I_T_ID
GET

ID_RO:= _ID;
END_GET
END_PROPERTY

PROPERTY PUBLIC Mode : KOSTAL_AF2024_Core_process.I_T_processMode
GET

Mode:= _mode;
END_GET
END_PROPERTY

PROPERTY PUBLIC Participants : I_ListOfParticipant
GET

Participants:= _Participants;
END_GET
END_PROPERTY

PROPERTY PUBLIC RunEmpty : BOOL
GET
RunEmpty := _runEmpty;
END_GET
END_PROPERTY

PROPERTY PUBLIC step : KOSTAL_AF2024_Core_process.I_processStep
GET

step:= _step;
END_GET
END_PROPERTY

END_FUNCTION_BLOCK

// Project Information/F_GetCompany
// This function has been automatically generated from the project information.
{attribute 'signature_flag' := '1073741824'}
{attribute 'TcGenerated'}
{attribute 'no-analysis'}
FUNCTION F_GetCompany : WSTRING
VAR_INPUT
	
END_VAR

F_GetCompany := "KOSTAL GmbH & Co.KG";

END_FUNCTION

// Project Information/F_GetTitle
// This function has been automatically generated from the project information.
{attribute 'signature_flag' := '1073741824'}
{attribute 'TcGenerated'}
{attribute 'no-analysis'}
FUNCTION F_GetTitle : WSTRING
VAR_INPUT
	
END_VAR

F_GetTitle := "KOSTAL.AF2024.Core.MainControl";

END_FUNCTION

// Project Information/F_GetVersion
// This function has been automatically generated from the project information.
{attribute 'signature_flag' := '1073741824'}
{attribute 'TcGenerated'}
{attribute 'no-analysis'}
FUNCTION F_GetVersion : ST_LibVersion
VAR_INPUT
	
END_VAR

F_GetVersion.iMajor := 1;
F_GetVersion.iMinor := 0;
F_GetVersion.iBuild := 0;
F_GetVersion.iRevision := 0;
F_GetVersion.sVersion := '1.0.0.0';
F_GetVersion.nFlags := 0;

END_FUNCTION
